Fanuc KAREL source: KO00146.KL

PROGRAM KO00146
%NOLOCKGROUP
VAR
  R: REAL
  CFG: CONFIG
  OUT: XYZWPR
  N: REAL
BEGIN
  N = 1
  R = 2.0
  CFG.CFG_FLIP = TRUE
  OUT = POS(R, R, R, R, N, R, CFG)
END KO00146
